(*
SPDX-FileCopyrightText: © 2026 Oleksandr Tiutyk <trofimich@gmail.com>
SPDX-License-Identifier: MIT
License: https://opensource.org/license/mit
*)

(*!
<summary>Stores the auto-dispose registry and fallback-cleanup diagnostics of one cyclic PLC task.</summary>
<description>
Internal manager storage. Only the owning task mutates it during cyclic execution. Application teardown may
release it after cyclic tasks have stopped. Objects belong to the registry; clients borrow references until
cleanup.
</description>
*)
TYPE TASK_MEMORY_STATE :
STRUCT
	Objects : POINTER TO IObject;
	BufferCapacity : DWORD;
	ObjectCount : DWORD;

	LastSystemTaskCycleCount : UDINT;
	MissedCleanupCount : UDINT;
END_STRUCT
END_TYPE

(* stored: Version 1.1.0.1
   DUT TASK_MEMORY_STATE: Id {53579067-3cc5-4a24-86a6-01cb0646981b} *)
